FUNCTION_BLOCK MainsSwitchbox (* CAT Function Block Type *)
  (* Standard: 61499-2 *)
  (* Version 0.0, 8/3/2026, template *)
  PACKAGE Main;
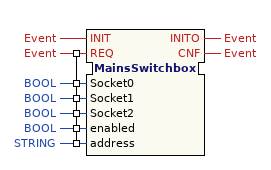
  EVENT_INPUT
    INIT; (* Initialization Request *)
    REQ WITH Socket0, Socket1, Socket2, enabled, address; (* Normal Execution Request *)
  END_EVENT
  EVENT_OUTPUT
    INITO; (* Initialization Confirm *)
    CNF; (* Execution Confirmation *)
  END_EVENT
  VAR_INPUT
    Socket0 : BOOL; (* Input event qualifier *)
    Socket1 : BOOL;
    Socket2 : BOOL;
    enabled : BOOL;
    address : STRING;
  END_VAR
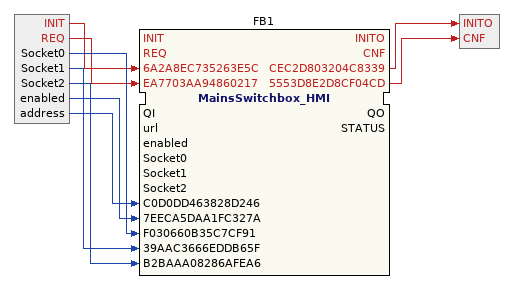
  FBS
    FB1 : MainsSwitchbox_HMI;
  END_FBS
  EVENT_CONNECTIONS
    INIT TO FB1.6A2A8EC735263E5C;
    REQ TO FB1.EA7703AA94860217;
    FB1.CEC2D803204C8339 TO INITO;
    FB1.5553D8E2D8CF04CD TO CNF;
  END_CONNECTIONS
  DATA_CONNECTIONS
    address TO FB1.C0D0DD463828D246;
    enabled TO FB1.7EECA5DAA1FC327A;
    Socket0 TO FB1.F030660B35C7CF91;
    Socket1 TO FB1.39AAC3666EDDB65F;
    Socket2 TO FB1.B2BAAA08286AFEA6;
  END_CONNECTIONS
END_FUNCTION_BLOCK
